(* IEC 61131-3 sources: PLC-Static-Analysis/modules/frontend-st/src/test/resources/golden, 24 files *)

(* ---- enum_trailing_comma.st ---- *)
// Enumerations with a comma after the last value (docs/grammar/codesys.md section 7, M12)
TYPE E_Handshake :
(
    Load := 1,
    CameraCheck := 2,
);
END_TYPE

TYPE E_SystemState :
(
    IDLE := 0,
    RUNNING := 1, // comment after the last comma
) WORD;
END_TYPE

TYPE E_Plain : (Red, Green, Blue,) := Green;
END_TYPE

(* ---- struct_qualifier.st ---- *)
// A qualifier after STRUCT applies to the whole structure (docs/grammar/codesys.md section 7, M12)
TYPE ST_Parameter :
STRUCT PERSISTENT
    rSetpoint : REAL := 1.5;
    nMode : INT;
END_STRUCT
END_TYPE

TYPE ST_AxisRetain :
STRUCT RETAIN
    lrPosition : LREAL;
END_STRUCT
END_TYPE

TYPE ST_Steps :
STRUCT CONSTANT
    nStart : INT := 10;
    nStop : INT := 20;
END_STRUCT
END_TYPE

(* ---- types.st ---- *)
TYPE
    ST_Point EXTENDS ST_Base :
    STRUCT
        x : REAL;
        y : REAL := 0.0;
    END_STRUCT
    E_State : (Idle := 0, Running, Faulted := 10) INT := Idle;
    U_Raw :
    UNION
        dw : DWORD;
        ab : ARRAY[0..3] OF BYTE;
    END_UNION
    T_Name : STRING(80);
    T_Percent : INT(0..100);
    T_Matrix : ARRAY[1..3, 1..3] OF LREAL;
    T_Ref : REF_TO INT;
END_TYPE

(* ---- pragmas_comments.st ---- *)
// line comment
(* outer (* nested *) still outer *)
/* C-style /* nested */ comment */
{attribute 'qualified_only'}
{attribute 'TcLinkTo' := '.in := TIIB[Term 1]^Channel 1^Value'}
VAR_GLOBAL
    {attribute 'pytmc' := '
        pv: TEST:VALUE
        io: i
    '}
    gValue : INT; // trailing comment
    {warning 'check this'}
    gOther : INT;
END_VAR
{IF defined (SIMULATION)}
{ELSE}
{END_IF}
{region "Main part"}
{endregion}

(* ---- error_exst_target.st ---- *)
// CODESYS ExST: the left side of an assignment in an expression must be a variable (M12)
FUNCTION F_Bad : BOOL
VAR
    a, b : BOOL;
END_VAR
IF (a AND b := TRUE) THEN
    F_Bad := TRUE;
END_IF
END_FUNCTION

(* ---- expressions.st ---- *)
FUNCTION F_Expr : LREAL
VAR_INPUT
    p : POINTER TO ST_Point;
END_VAR
VAR
    w : WORD;
    s : STRING;
    ws : WSTRING;
    b : BOOL;
    t : TIME;
END_VAR

F_Expr := -2 ** 2 + 3 * 4 MOD 5 - (1 + 2) / 3;
b := NOT b AND w.3 OR_ELSE p^.x > 1.5E-3 AND_THEN THIS^.bOk XOR SUPER^.bOk;
b := 1 < 2 = TRUE <> FALSE;
w := 16#FF_FF + 2#1010 + 8#17 + 10#99 + WORD#16#0F + INT#-5;
s := 'it$'s $N done';
ws := "wide $"quoted$"";
t := T#1h2m3s4ms + LTIME#-5us;
F_Expr := TO_LREAL(D#2024-01-31 - DATE#2024-01-01) + TOD#12:30:15.5 + DT#2024-01-31-12:00:00;
w := SIZEOF(POINTER TO ST_Point) + SIZEOF(STRING) + .gGlobal + AND(b, b);
F_Expr := arr[i, j + 1].field;
END_FUNCTION

(* ---- config_oop.st ---- *)
NAMESPACE Lib.Motion
USING Lib.Base, Other;
INTERFACE I_Axis EXTENDS I_Base, I_Diag
METHOD MoveAbs : BOOL
VAR_INPUT
    pos : LREAL;
END_VAR
END_METHOD
PROPERTY Position : LREAL
END_PROPERTY
END_INTERFACE
CLASS FINAL C_Axis IMPLEMENTS I_Axis
VAR PUBLIC
    pos : LREAL;
END_VAR
METHOD PUBLIC OVERRIDE MoveAbs : BOOL
MoveAbs := TRUE;
END_METHOD
END_CLASS
END_NAMESPACE

CONFIGURATION Cfg
VAR_GLOBAL
    gRun : BOOL;
END_VAR
RESOURCE Res ON PLC
    TASK Fast(INTERVAL := T#10MS, PRIORITY := 1);
    PROGRAM Main WITH Fast : MAIN;
END_RESOURCE
END_CONFIGURATION

(* ---- error_misplaced_implements.st ---- *)
FUNCTION_BLOCK FB_A
VAR
    x : INT;
END_VAR
IMPLEMENTS I_A
x := 1;
END_FUNCTION_BLOCK

FUNCTION_BLOCK FB_B
VAR_GENERIC CONSTANT
    n : INT := 1;
END_VAR
VAR
    y : INT;
END_VAR
EXTENDS FB_A
END_FUNCTION_BLOCK

PROGRAM P
VAR_GENERIC CONSTANT
    n : INT := 1;
END_VAR
IMPLEMENTS I_A
END_PROGRAM

(* ---- error_missing_operand.st ---- *)
FUNCTION_BLOCK FB_Template
VAR
    eState : E_PROGRESS;
    nErrorId : UDINT;
    fbMove : FB_Move;
END_VAR
// Unfinished template code (pattern from a vendor XTS demo): each mistake should give one diagnostic.
IF fbMove.Error THEN
    eState := E_PROGRESS.PROGRESS_ERROR;
    nErrorId :=

ELSIF fbMove.Done THEN
    eState := E_PROGRESS.;

END_IF
CASE eState OF
    E_PROGRESS.PROGRESS_BUSY:
        nErrorId := nErrorId *;
END_CASE
nErrorId := fbMove.;
eState := E_PROGRESS.PROGRESS_INIT;
END_FUNCTION_BLOCK

(* ---- exst_assignment_expression.st ---- *)
// CODESYS ExST: an assignment used as an expression (docs/grammar/codesys.md section 7, M12)
FUNCTION_BLOCK FB_ExSt
VAR
    b, bInit, bOk : BOOL;
    i, n : INT;
    s : STRING;
    p : POINTER TO INT;
    st : ST_Item;
    arr : ARRAY[0..9] OF INT;
END_VAR

// whole condition: the value is the rest of the expression
IF b := (i = 1) THEN
    i := i + 1;
ELSIF st.bDone := i > 2 OR b THEN
    i := 0;
END_IF
WHILE p^ := p^ - 1 DO
    ;
END_WHILE
REPEAT
    i := i + 1;
UNTIL bOk := i >= 10
END_REPEAT

// in parentheses, anywhere an expression is
IF (n := FIND(s, 'x')) > 0 AND_THEN (arr[n] := n * 2) <> 0 THEN
    s := '';
END_IF
CASE (n := n + 1) OF
    1: i := 1;
END_CASE
b := NOT (bOk := fbChild.Execute());
RETURN(bInit := i <= 0);

// statement level stays a chained assignment
i := n := 0;
END_FUNCTION_BLOCK

(* ---- generic_fb.st ---- *)
(* Generic function blocks (CODESYS help "VAR_GENERIC CONSTANT"): generic constants come before EXTENDS / IMPLEMENTS *)
FUNCTION_BLOCK FB_MyString
VAR_GENERIC CONSTANT
    maxlen : UDINT := 1;
END_VAR
IMPLEMENTS IString, IPrintable
VAR
    buffer : ARRAY[0..maxlen] OF BYTE;
END_VAR
buffer[0] := 0;
END_FUNCTION_BLOCK

FUNCTION_BLOCK FB_MySpecialString
VAR_GENERIC CONSTANT
    maxlen2 : UDINT := 1;
END_VAR
EXTENDS FB_MyString<maxlen2> IMPLEMENTS ISpecial
END_FUNCTION_BLOCK

FUNCTION_BLOCK FB_LongString EXTENDS FB_MyString<1000>
END_FUNCTION_BLOCK

PROGRAM MAIN
VAR
    s : FB_MyString<(2 * 5)>;
END_VAR
s();
END_PROGRAM

(* ---- il_pous.st ---- *)
(* Instruction List POUs next to an ST one *)
FUNCTION_BLOCK FB_Distance
VAR_INPUT
    X1, X2, Y1, Y2 : REAL;
    TMax : REAL;
END_VAR
VAR_OUTPUT
    Dist : REAL;
    Ok : BOOL;
END_VAR
VAR
    Temp : REAL;
    Pulse : TON;
END_VAR
    LD   Y1
    SUB  Y2         (* Y1 - Y2 *)
    ST   Temp
    MUL  Temp
    ADD( X1         (* deferred: + (X1 - X2)^2 *)
    SUB  X2
    ST   Temp
    MUL  Temp
    )
    SQRT
    ST   Dist
    GT   TMax
    JMPC TooFar
    S    Ok
    CAL  Pulse(IN := Ok,
               PT := T#1S)
    RET
TooFar:
    LDN  Pulse.Q
    R    Ok
END_FUNCTION_BLOCK

PROGRAM Counter
VAR
    Count : INT;
    Done : BOOL;
END_VAR
LD Count;
ADD 1;
ST Count;
GE 10;
ST Done;
END_PROGRAM

FUNCTION_BLOCK FB_St
VAR
    a : INT;
END_VAR
a := a + 1;
END_FUNCTION_BLOCK

(* ---- keyword_names.st ---- *)
(* CONTINUE as a variable name: declared, read, written, as a member; CONTINUE; stays the loop statement. *)
FUNCTION_BLOCK FB_Axis
VAR_INPUT
    Power : BOOL;
    SingleStep : BOOL;
    Continue : BOOL;
    MoveInterrupted : BOOL;
END_VAR
VAR
    i : INT;
END_VAR
IF Continue THEN
    Continue := FALSE;
END_IF
FOR i := 1 TO 10 DO
    IF i = 5 THEN
        CONTINUE;
    END_IF
END_FOR
END_FUNCTION_BLOCK

PROGRAM MAIN
VAR
    fbMy6Axis : FB_Axis;
    bEnable : BOOL;
END_VAR
IF fbMy6Axis.Power=TRUE AND fbMy6Axis.SingleStep=TRUE THEN
    IF fbMy6Axis.Continue=TRUE AND fbMy6Axis.MoveInterrupted=TRUE THEN
        fbMy6Axis.Continue:=FALSE;
    END_IF
    fbMy6Axis(Continue := bEnable);
END_IF
END_PROGRAM

(* ---- missing_semicolon_accepted.st ---- *)
// A ';' left out before END_VAR or after the last statement of a body: a warning (docs/grammar/codesys.md, M12)
FUNCTION_BLOCK FB_Collection
VAR_INPUT
    bInitRetains : BOOL; // initialise retain variables
    T : Tc2_Utilities.T_Arg // provide the type of the collection
END_VAR
VAR_IN_OUT
    XTSUnitRef : I_XtsUnit//FB_XtsUnit;
END_VAR
VAR
    n : INT;
END_VAR
n := n + 1;
Engine.oRun := n > 2
METHOD M : BOOL
M := TRUE
END_METHOD
END_FUNCTION_BLOCK

FUNCTION F_Speed : UINT
VAR_INPUT
    iAnalog : INT;
END_VAR
F_Speed := TO_UINT(LIMIT(0, iAnalog, 24000))

(* ---- pou_function_block.st ---- *)
(* Function block with inheritance, all variable sections, methods, a property and an action. *)
{attribute 'reflection'}
FUNCTION_BLOCK PUBLIC FB_Motor EXTENDS FB_Base IMPLEMENTS I_Motor, I_Diag
VAR_INPUT
    bStart : BOOL;
    rSetpoint : REAL := 1.5;
END_VAR
VAR_OUTPUT
    bRunning AT %QX0.1 : BOOL;
END_VAR
VAR_IN_OUT
    stConfig : ST_Config;
END_VAR
VAR RETAIN PERSISTENT
    nStarts : UDINT;
END_VAR
VAR CONSTANT
    MAX_SPEED : INT := 1500;
END_VAR
VAR
    {attribute 'hide'}
    fbTimer : TON := (PT := T#2S);
    aBuf : ARRAY[0..9] OF INT := [1, 2, 8(0)];
    pData : POINTER TO BYTE;
    refCfg : REFERENCE TO ST_Config;
    fbInit : FB_Logger(10, sName := 'motor');
    a, b : INT;
END_VAR

fbTimer(IN := bStart, Q => bRunning);
IF bRunning THEN
    nStarts := nStarts + 1;
END_IF

METHOD PUBLIC Reset : BOOL
VAR_INPUT
    bForce : BOOL;
END_VAR
nStarts := 0;
Reset := TRUE;
END_METHOD

PROPERTY PUBLIC Speed : INT
GET
    Speed := MAX_SPEED;
END_GET
SET
    ;
END_SET
END_PROPERTY

ACTION Stop:
    bRunning := FALSE;
END_ACTION
END_FUNCTION_BLOCK

(* ---- text_export_no_end.st ---- *)
FUNCTION_BLOCK FB_Exported
VAR_INPUT
    bIn : BOOL;
END_VAR
VAR
    n : INT;
END_VAR
IF bIn THEN
    n := n + 1;
END_IF

(* ---- array_init_no_brackets.st ---- *)
// Array initial values without brackets, CODESYS V2 style (docs/grammar/codesys.md section 7, M12)
PROGRAM P
VAR
    buf : ARRAY[0..3] OF BYTE := 110, 60, 3, 219; (* crypt key *)
    arr2 : ARRAY[1..2, 3..4] OF INT := 1, 3(7);
    arr3 : ARRAY[1..8] OF INT := 2(0), 4(4), 2, 3;
    one : ARRAY[1..3] OF INT := 3(5);
    n : INT := 5;
END_VAR
n := n + 1;
END_PROGRAM

(* ---- error_missing_semicolon.st ---- *)
// A ';' left out anywhere else stays a syntax error (docs/grammar/codesys.md, M12)
TYPE ST_Row :
STRUCT
    a : INT;
    b : BOOL
END_STRUCT
END_TYPE

PROGRAM P
VAR
    a : INT
    b : INT;
END_VAR
a := 1
b := 2;
IF a > 0 THEN
    b := 3
END_IF
CASE a OF
    1: b := 4
    2: b := 5;
END_CASE
END_PROGRAM

(* ---- error_recovery.st ---- *)
PROGRAM P
VAR
    a : INT;
    b : INT := ;
    c : BOOL;
END_VAR
a := 1 +;
c := TRUE;
IF a > 1 THEN
    a := 2
END_IF
a FOO= 3;
§
c := FALSE;
b := 'unterminated
END_PROGRAM

(* ---- error_unterminated_comment.st ---- *)
PROGRAM P
VAR a : INT; END_VAR
a := 1;
(* this comment (* nests *) and is never closed
a := 2;

(* ---- repeat_count_expression.st ---- *)
// Array repetition counts that are constant expressions (docs/grammar/codesys.md section 7, M12)
VAR_GLOBAL CONSTANT
    N : INT := 4;
END_VAR

PROGRAM P
VAR
    aText : ARRAY[0..N] OF STRING(255) := [N + 1(',')];
    aFlags : ARRAY[0..N - 1] OF ST_Flag := [(N - 1)((bOn := TRUE, sName := '')), (bOn := FALSE, sName := 'x')];
    aMix : ARRAY[1..6] OF INT := [2(0), GVL.M(1), 3];
    aCalls : ARRAY[1..2] OF INT := [F(1), F(2)];
END_VAR
aText[0] := '';
END_PROGRAM

(* ---- statements.st ---- *)
PROGRAM MAIN
VAR
    i, n : INT;
    eState : E_State;
    bA, bB, bC : BOOL;
    r : REFERENCE TO INT;
    itf : I_Motor;
END_VAR

CASE eState OF
    E_State.Idle, E_State#Running:
        n := 1;
    1..5, 7:
        n := 2;
ELSE
    n := 0;
END_CASE;

FOR i := 0 TO 10 BY 2 DO
    IF i = 4 THEN CONTINUE; END_IF
    IF i > 8 THEN EXIT; END_IF
END_FOR

WHILE n < 10 DO n := n + 1; END_WHILE
REPEAT n := n - 1; UNTIL n <= 0 END_REPEAT

bA S= bB;
bA R= bC;
r REF= n;
itf ?= fbAny;
bA := bB := bC := FALSE;

JMP lbl;
lbl:
__TRY
    n := 1 / n;
__CATCH(exc)
    n := 0;
__FINALLY
    ;
__ENDTRY

fbT(IN := bA, PT := T#1S, Q => bB, NOT ET => );
RETURN;
END_PROGRAM

(* ---- statements_only.st ---- *)
// an exported action body: statements without any declaration
nCount := nCount + 1;
IF nCount > 10 THEN
    nCount := 0;
END_IF

(* ---- type_modifier_empty_init.st ---- *)
// TYPE with an access modifier, empty structured initialisers (docs/grammar/codesys.md section 7, M12)
TYPE INTERNAL E_State :
(
    Idle,
    Busy
);
END_TYPE

TYPE INTERNAL ST_Row :
STRUCT
    a : INT;
    b : BOOL;
END_STRUCT
END_TYPE

PROGRAM P
VAR
    fbList : FB_List := ();
    stRow : ST_Row := ();
    fbFree : FB_Free(42) := ();
    aRows : ARRAY[1..15] OF ST_Row := [15(())];
    aMixed : ARRAY[1..3] OF ST_Row := [(a := 1), 2(())];
END_VAR
stRow.a := 1;
END_PROGRAM
